(* IEC 61131-3 sources: SRCI_CLIENT_PLC/RobotLibrary/Library/POUs/Write/MC_WriteToolData/Structures, 4 files *)

(* ---- WriteToolDataOutCmd.st ---- *)
{attribute 'pack_mode' := '1'}
// -------------------------------------------------------------------------
//  SRCI Robot Library
// -------------------------------------------------------------------------
//
//  Object:      WriteToolDataOutCmd
//  Author:      Thorsten Brach
//  Date:        2024-08-08
//
//  Description:
//
//
//  Copyright:
//    (C) 2024 Thorsten Brach. All rights reserved
//             Licensed under the MIT License.
//
//  Disclaimer:
//    This project is provided without any guarantee and can be used for
//    private and commercial purposes. Any use is at the user’s
//    own risk and responsibility.
//
// -------------------------------------------------------------------------
TYPE WriteToolDataOutCmd :
STRUCT
END_STRUCT
END_TYPE

(* ---- WriteToolDataParCmd.st ---- *)
{attribute 'pack_mode' := '1'}
// -------------------------------------------------------------------------
//  SRCI Robot Library
// -------------------------------------------------------------------------
//
//  Object:      WriteToolDataParCmd
//  Author:      Thorsten Brach
//  Date:        2024-08-08
//
//  Description:
//
//
//  Copyright:
//    (C) 2024 Thorsten Brach. All rights reserved
//             Licensed under the MIT License.
//
//  Disclaimer:
//    This project is provided without any guarantee and can be used for
//    private and commercial purposes. Any use is at the user’s
//    own risk and responsibility.
//
// -------------------------------------------------------------------------
TYPE WriteToolDataParCmd :
STRUCT
  /// Tool index
  /// •      0: Flange (default) Not possible to change
  /// • 1..254: Tool Frame
  ToolNo            : USINT;
  /// Tool data (see chapter 5.5.6.3)
  ToolData          : ToolData;
END_STRUCT
END_TYPE

(* ---- WriteToolDataRecvData.st ---- *)
{attribute 'pack_mode' := '1'}
// -------------------------------------------------------------------------
//  SRCI Robot Library
// -------------------------------------------------------------------------
//
//  Object:      WriteToolDataRecvData
//  Author:      Thorsten Brach
//  Date:        2024-08-08
//
//  Description:
//
//
//  Copyright:
//    (C) 2024 Thorsten Brach. All rights reserved
//             Licensed under the MIT License.
//
//  Disclaimer:
//    This project is provided without any guarantee and can be used for
//    private and commercial purposes. Any use is at the user’s
//    own risk and responsibility.
//
// -------------------------------------------------------------------------
TYPE WriteToolDataRecvData EXTENDS RspHeader :
STRUCT
END_STRUCT
END_TYPE

(* ---- WriteToolDataSendData.st ---- *)
{attribute 'pack_mode' := '1'}
// -------------------------------------------------------------------------
//  SRCI Robot Library
// -------------------------------------------------------------------------
//
//  Object:      WriteToolDataSendData
//  Author:      Thorsten Brach
//  Date:        2024-08-08
//
//  Description:
//
//
//  Copyright:
//    (C) 2024 Thorsten Brach. All rights reserved
//             Licensed under the MIT License.
//
//  Disclaimer:
//    This project is provided without any guarantee and can be used for
//    private and commercial purposes. Any use is at the user’s
//    own risk and responsibility.
//
// -------------------------------------------------------------------------
TYPE WriteToolDataSendData EXTENDS CmdHeader:
STRUCT
  /// Reserve
  Reserve           : BYTE;
  /// Tool index
  /// •      0: Flange (default) Not possible to change
  /// • 1..254: Tool Frame
  ToolNo            : USINT;
  /// Tool data (see chapter 5.5.6.3)
  ToolData          : ToolData;
END_STRUCT
END_TYPE
